FUNCTION_BLOCK Algorithm_p (* Basic Function Block Type *)
  (* Standard: 61499-2 *)
  (* Version 0.0, 10/22/2026, macie, Schneider Electric, Template *)
  PACKAGE Main;
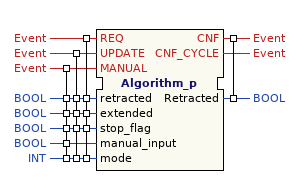
  EVENT_INPUT
    REQ WITH retracted, extended, stop_flag, mode; (* Normal Execution Request *)
    UPDATE WITH retracted, extended, stop_flag, mode;
    MANUAL WITH retracted, extended, stop_flag, manual_input, mode;
  END_EVENT
  EVENT_OUTPUT
    CNF WITH Retracted; (* Execution Confirmation *)
    CNF_CYCLE;
  END_EVENT
  VAR_INPUT
    retracted : BOOL; (* Input event qualifier *)
    extended : BOOL;
    stop_flag : BOOL;
    manual_input : BOOL;
    mode : INT;
  END_VAR
  VAR_OUTPUT
    Retracted : BOOL; (* Output event qualifier *)
  END_VAR
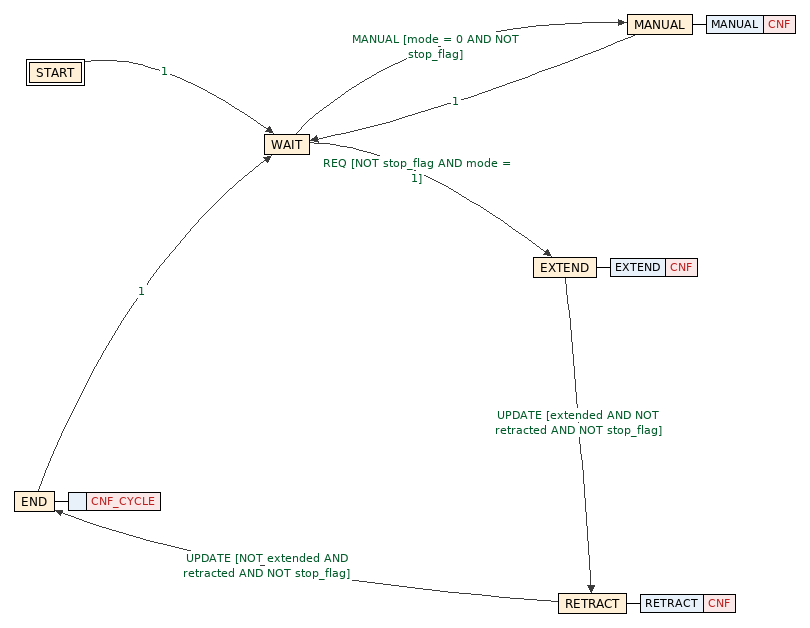
  EC_STATES
    START; (* Initial State *)
    WAIT;
    EXTEND : EXTEND -> CNF;
    RETRACT : RETRACT -> CNF;
    END : -> CNF_CYCLE;
    MANUAL : MANUAL -> CNF;
  END_STATES
  EC_TRANSITIONS
    WAIT TO EXTEND := REQ [NOT stop_flag AND mode = 1];
    START TO WAIT := 1;
    EXTEND TO RETRACT := UPDATE [extended AND NOT retracted AND NOT stop_flag];
    RETRACT TO END := UPDATE [NOT extended AND retracted AND NOT stop_flag];
    END TO WAIT := 1;
    WAIT TO MANUAL := MANUAL [mode = 0 AND NOT stop_flag];
    MANUAL TO WAIT := 1;
  END_TRANSITIONS
  ALGORITHM RETRACT IN ST: (* Initialization algorithm *)
;
Retracted := FALSE;
  END_ALGORITHM
  ALGORITHM EXTEND IN ST: (* Normally executed algorithm *)
;
Retracted := TRUE;
  END_ALGORITHM
  ALGORITHM MANUAL IN ST:
;
Retracted := manual_input;
  END_ALGORITHM
END_FUNCTION_BLOCK
